FUNCTION_BLOCK Controller (* Composite Function Block Type *)
  (* Standard: 61499-2 *)
  (* Version 0.0, 7/13/2016, Andrei, nxtControl GmbH, template *)
  PACKAGE Main;
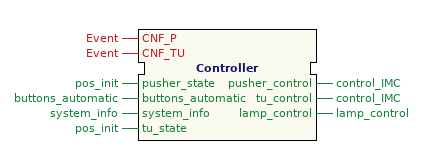
  EVENT_INPUT
    CNF_P;
    CNF_TU;
  END_EVENT
  SOCKETS
    pusher_state : pos_init;
    buttons_automatic : buttons_automatic;
    system_info : system_info;
    tu_state : pos_init;
  END_SOCKETS
  PLUGS
    pusher_control : control_IMC;
    tu_control : control_IMC;
    lamp_control : lamp_control;
  END_PLUGS
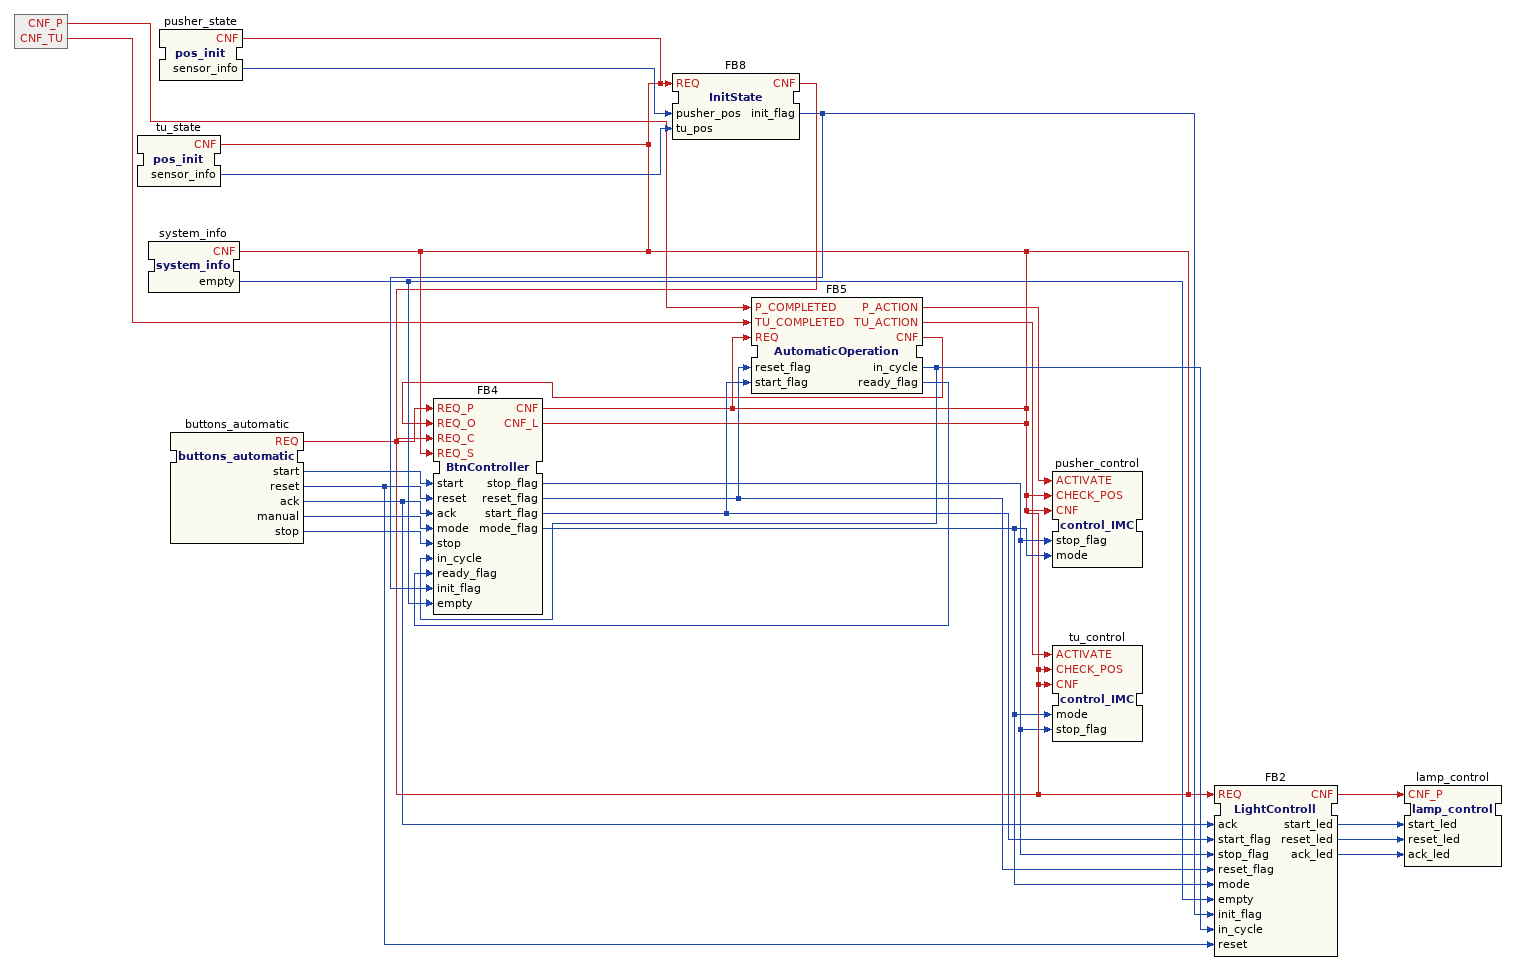
  FBS
    FB4 : BtnController;
    FB5 : AutomaticOperation;
    FB2 : LightControll;
    FB8 : InitState;
  END_FBS
  EVENT_CONNECTIONS
    FB8.CNF TO FB4.REQ_C;
    FB4.CNF_L TO FB2.REQ;
    pusher_state.CNF TO FB8.REQ;
    buttons_automatic.REQ TO FB4.REQ_P;
    buttons_automatic.REQ TO FB2.REQ;
    system_info.CNF TO FB8.REQ;
    system_info.CNF TO FB2.REQ;
    FB2.CNF TO lamp_control.CNF_P;
    tu_state.CNF TO FB8.REQ;
    CNF_P TO FB5.P_COMPLETED;
    CNF_TU TO FB5.TU_COMPLETED;
    FB5.CNF TO FB4.REQ_O;
    FB5.P_ACTION TO pusher_control.ACTIVATE;
    FB5.TU_ACTION TO tu_control.ACTIVATE;
    system_info.CNF TO pusher_control.CHECK_POS;
    system_info.CNF TO tu_control.CHECK_POS;
    FB4.CNF TO FB5.REQ;
    FB4.CNF TO pusher_control.CNF;
    FB4.CNF TO tu_control.CNF;
    system_info.CNF TO FB4.REQ_S;
    FB4.CNF TO FB2.REQ;
  END_CONNECTIONS
  DATA_CONNECTIONS
    FB4.reset_flag TO FB5.reset_flag;
    FB4.start_flag TO FB5.start_flag;
    FB4.stop_flag TO FB2.stop_flag;
    FB4.start_flag TO FB2.start_flag;
    FB4.reset_flag TO FB2.reset_flag;
    FB4.mode_flag TO FB2.mode;
    FB5.in_cycle TO FB4.in_cycle;
    FB8.init_flag TO FB4.init_flag;
    FB8.init_flag TO FB2.init_flag;
    FB5.in_cycle TO FB2.in_cycle;
    pusher_state.sensor_info TO FB8.pusher_pos;
    FB4.stop_flag TO pusher_control.stop_flag;
    buttons_automatic.start TO FB4.start;
    buttons_automatic.reset TO FB4.reset;
    buttons_automatic.ack TO FB4.ack;
    buttons_automatic.manual TO FB4.mode;
    buttons_automatic.stop TO FB4.stop;
    buttons_automatic.reset TO FB2.reset;
    buttons_automatic.ack TO FB2.ack;
    system_info.empty TO FB2.empty;
    FB4.mode_flag TO pusher_control.mode;
    FB2.start_led TO lamp_control.start_led;
    FB2.reset_led TO lamp_control.reset_led;
    FB2.ack_led TO lamp_control.ack_led;
    FB4.mode_flag TO tu_control.mode;
    FB4.stop_flag TO tu_control.stop_flag;
    tu_state.sensor_info TO FB8.tu_pos;
    FB5.ready_flag TO FB4.ready_flag;
    system_info.empty TO FB4.empty;
  END_CONNECTIONS
END_FUNCTION_BLOCK
